TYPE ST_Recipe :
STRUCT
	rTargetKg   : LREAL;
	rBulkCutoff : LREAL := 0.9;
	sName       : STRING(40);
END_STRUCT
END_TYPE

(* stored: Version 1.1.0.1, ProductVersion 3.1.4024.12
   DUT ST_Recipe: Id {aaaaaaaa-0000-0000-0000-000000000008} *)
